// Règle de remise à zéro d'une variable de mover (docs/05 § 5.8)
{attribute 'qualified_only'}
{attribute 'strict'}
TYPE E_MoverVarReset :
(
    Never := 0,
    OnDeploy := 1,
    OnEmpty := 2
) USINT;
END_TYPE

(* stored: Version 1.1.0.1, ProductVersion 3.1.4024.12
   DUT E_MoverVarReset: Id {f339475a-bf5c-5137-a23e-a5c03e5e6e0b} *)
